(* LS Electric XG5000 project: NewProject *)
(* PLC LSPLC *)

PROGRAM NewProgram (* task: 스캔 프로그램 *)
VAR
    FF : FF;
END_VAR

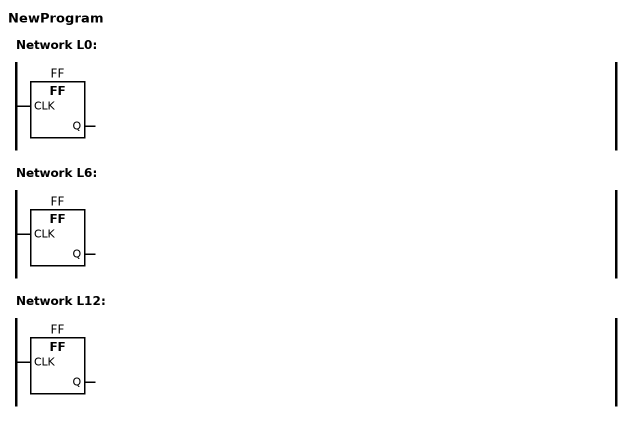
(* Rung L0 *)
FF(CLK := TRUE);
(* Rung L6 *)
FF(CLK := TRUE);
(* Rung L12 *)
FF(CLK := TRUE);
END_PROGRAM